(* IEC 61131-3 sources: SortJet_MasterSPS_Aufbau.fbsproj/08_POUs/Basis Funktionen/Switch Funktionen, 8 files *)

(* ---- LowHighByteSwitchInDWORD_CompleteSwap.fn.st ---- *)
(* METADATA
{
	"v3Meta": {
		"objectGuid": "8525d255-55de-4882-b974-c7e29f794d79"
	}
}
*)
FUNCTION LowHighByteSwitchInDWORD_CompleteSwap : DWORD
VAR_INPUT

  dwInputWord : DWORD;

END_VAR
VAR

  dwByte1 : DWORD;
  dwByte2 : DWORD;
  dwByte3 : DWORD;
  dwByte4 : DWORD;

END_VAR
dwByte1 :=SHR(dwInputWord,24);

dwByte2  :=SHL(dwInputWord,8);
dwByte2  :=SHR(dwByte2,24);
dwByte2  :=SHL(dwByte2,8);

dwByte3  :=SHL(dwInputWord,16);
dwByte3  :=SHR(dwByte3,24);
dwByte3  :=SHL(dwByte3,16);

dwByte4  :=SHL(dwInputWord,24);

LowHighByteSwitchInDWORD_CompleteSwap := dwByte1 OR dwByte2 OR dwByte3 OR dwByte4;
END_FUNCTION

(* ---- SWAP_DINT.fn.st ---- *)
(* METADATA
{
	"v3Meta": {
		"objectGuid": "60b6ea4b-319e-4cbc-b276-a980379624c0"
	}
}
*)
FUNCTION SWAP_DINT : DINT
VAR_INPUT

  // REAL
  dipWert : DINT;

END_VAR

VAR

  // BYTE
  aInByte  : ARRAY [0..3] OF BYTE ;
  aOutByte : ARRAY [0..3] OF BYTE ;

END_VAR
SysMemCpy( ADR(aInByte), ADR(dipWert),4 );

aOutByte[0] := aInByte[2];
aOutByte[1] := aInByte[3];
aOutByte[2] := aInByte[0];
aOutByte[3] := aInByte[1];

SysMemCpy( ADR(SWAP_DINT), ADR(aOutByte),4 );
END_FUNCTION

(* ---- SWAP_DWORD.fn.st ---- *)
(* METADATA
{
	"v3Meta": {
		"objectGuid": "389b713c-1c94-40ba-a43c-d7e5339b8bcd"
	}
}
*)
FUNCTION SWAP_DWORD : DWORD
VAR_INPUT

  // REAL
  dwpWert : DWORD;

END_VAR

VAR

  // BYTE
  aInByte  : ARRAY [0..3] OF BYTE ;
  aOutByte : ARRAY [0..3] OF BYTE ;

END_VAR
SysMemCpy( ADR(aInByte), ADR(dwpWert),4 );

aOutByte[0] := aInByte[3];
aOutByte[1] := aInByte[2];
aOutByte[2] := aInByte[1];
aOutByte[3] := aInByte[0];

SysMemCpy( ADR(SWAP_DWORD), ADR(aOutByte),4 );
END_FUNCTION

(* ---- SWAP_DWORD_SIEMENS.fn.st ---- *)
(* METADATA
{
	"v3Meta": {
		"objectGuid": "2a9c4065-11ba-4ec5-a5c1-2bac7310293a"
	}
}
*)
FUNCTION SWAP_DWORD_SIEMENS : DWORD
VAR_INPUT

  // REAL
  dwpWert : DWORD;

END_VAR

VAR

  // BYTE
  aInByte  : ARRAY [0..3] OF BYTE ;
  aOutByte : ARRAY [0..3] OF BYTE ;

END_VAR
SysMemCpy( ADR(aInByte), ADR(dwpWert),4 );

aOutByte[0] := aInByte[1];
aOutByte[1] := aInByte[0];
aOutByte[2] := aInByte[3];
aOutByte[3] := aInByte[2];

SysMemCpy( ADR(SWAP_DWORD_SIEMENS), ADR(aOutByte),4 );
END_FUNCTION

(* ---- SWAP_LOW_HIGH_WORD.fn.st ---- *)
(* METADATA
{
	"v3Meta": {
		"objectGuid": "88f4a337-90ad-4f2e-9ea2-c1124a4e2a48"
	}
}
*)
FUNCTION SWAP_LOW_HIGH_WORD : DWORD
VAR_INPUT
  IN : DWORD;
END_VAR
VAR
END_VAR
(* Hinweis:
   - Diese Funktion tauscht das LOW-WORD und das HIGH- WORD;
*)
SWAP_LOW_HIGH_WORD := ROL(IN, 16);
END_FUNCTION

(* ---- SWAP_REAL.fn.st ---- *)
(* METADATA
{
	"v3Meta": {
		"objectGuid": "ba889dae-5568-4c09-9bf3-2bdc011b0f01"
	}
}
*)
FUNCTION SWAP_REAL : REAL
VAR_INPUT

  // REAL
  rpWert : REAL;

END_VAR

VAR

  // BYTE
  aInByte  : ARRAY [0..3] OF BYTE ;
  aOutByte : ARRAY [0..3] OF BYTE ;

END_VAR
SysMemCpy( ADR(aInByte), ADR(rpWert),4 );

//aOutByte[0] := aInByte[3];
//aOutByte[1] := aInByte[2];
//aOutByte[2] := aInByte[1];
//aOutByte[3] := aInByte[0];

aOutByte[0] := aInByte[1];
aOutByte[1] := aInByte[0];
aOutByte[2] := aInByte[3];
aOutByte[3] := aInByte[2];

SysMemCpy( ADR(SWAP_REAL), ADR(aOutByte),4 );
END_FUNCTION

(* ---- SWAP_REAL_SIEMENS.fn.st ---- *)
(* METADATA
{
	"v3Meta": {
		"objectGuid": "24a74364-fccd-4a66-8b87-fbfc150829ad"
	}
}
*)
FUNCTION SWAP_REAL_SIEMENS : REAL
VAR_INPUT

  // REAL
  rpWert : REAL;

END_VAR

VAR

  // BYTE
  aInByte  : ARRAY [0..3] OF BYTE ;
  aOutByte : ARRAY [0..3] OF BYTE ;

END_VAR
SysMemCpy( ADR(aInByte), ADR(rpWert),4 );

aOutByte[0] := aInByte[2];
aOutByte[1] := aInByte[3];
aOutByte[2] := aInByte[0];
aOutByte[3] := aInByte[1];
SysMemCpy( ADR(SWAP_REAL_SIEMENS), ADR(aOutByte),4 );
END_FUNCTION

(* ---- SWAP_WORD.fn.st ---- *)
(* METADATA
{
	"v3Meta": {
		"objectGuid": "f5bf0334-c8db-496d-a0a5-3bfc853a0111"
	}
}
*)
FUNCTION SWAP_WORD : WORD
VAR_INPUT

  // BOOELAN
  wpWert : WORD;

END_VAR
VAR

  // BYTE
  aInByte  : ARRAY [0..1] OF BYTE ;
  aOutByte : ARRAY [0..1] OF BYTE ;

END_VAR
SysMemCpy( ADR(aInByte), ADR(wpWert),2 );

aOutByte[0] := aInByte[1];
aOutByte[1] := aInByte[0];

SysMemCpy( ADR(SWAP_WORD), ADR(aOutByte),2 );
END_FUNCTION
